(* IEC 61131-3 sources: SortJet_MasterSPS_Aufbau.fbsproj/Device.device.xml.v3^/Plc Logic.plclogic.xml.v3^/Application.application.xml.v3^/00_Basis/StationBasisZuweisungen.prg.st^, 20 files *)

(* ---- M_AufrufeZuweisungen.meth.st ---- *)
(* METADATA
{
	"v3Meta": {
		"objectGuid": "6343c508-4884-483e-a331-d4339a485652"
	}
}
*)
METHOD M_AufrufeZuweisungen
VAR_INPUT
END_VAR
VAR
  wlIndex : WORD;
END_VAR

//-------------------------------------------------------------------------------------------------
// PARAMETER ZUWEISEN
//-------------------------------------------------------------------------------------------------

// Aufrufe der Zuweisungen
Zuweisung_101();
Zuweisung_102();
Zuweisung_151();
Zuweisung_152();
Zuweisung_201();
Zuweisung_202();
Zuweisung_203();
Zuweisung_204();
Zuweisung_205();
Zuweisung_206();
Zuweisung_207();
Zuweisung_208();

Zuweisung_301();
Zuweisung_302();
Zuweisung_303();
Zuweisung_304();
Zuweisung_305();

Zuweisung_401();

Zuweisung_501();
END_METHOD

(* ---- Zuweisung_101.act.st ---- *)
(* METADATA
{
	"v3Meta": {
		"objectGuid": "51c9bc00-b1a7-48c3-ab96-ac2ea4b83acf"
	}
}
*)
ACTION Zuweisung_101
// Zuweisung der MK's
starrShuttleBasisParameter[cSHUTTLE_101].stMKs REF= apgMKShuttle101;

// Antriebsparameter zuweisen
starrShuttleBasisParameter[cSHUTTLE_101].stAntriebsparameter.stGlastransport                   REF= apgInfoShuttle101Glastransport;
starrShuttleBasisParameter[cSHUTTLE_101].stAntriebsparameter.stGlastransportSlave              REF= apgInfoShuttle101GlastransportSlave;
starrShuttleBasisParameter[cSHUTTLE_101].stAntriebsparameter.stWandverstellung                 REF= apgInfoShuttle101Dickenverstellung;
starrShuttleBasisParameter[cSHUTTLE_101].stParameterStationskomponenten.stGlastransportShuttle REF= apgMKShuttle101Glastransport;
starrShuttleBasisParameter[cSHUTTLE_101].stParameterStationskomponenten.stKippen               REF= apgMKShuttle101Kippen;
starrShuttleBasisParameter[cSHUTTLE_101].stParameterStationskomponenten.stWandverstellung      REF= apgMKShutte101Scheibenfuehrung;

starrShuttleBasisParameter[cSHUTTLE_101].stAntriebsparameter.stQuerfahrt REF= apgInfoShuttle101Querfahrt;
starrShuttleBasisParameter[cSHUTTLE_101].stAntriebsparameter.stKippen    REF= apgInfoShuttle101Kippen;

// Greifer [Ausbaustufe stStationsAufbau.bGreifer]
starrShuttleBasisParameter[cSHUTTLE_101].stParameterStationskomponenten.stGreifer REF= apgMKShuttle101Greifer;
starrShuttleBasisParameter[cSHUTTLE_101].stAntriebsparameter.stGreifer            REF= apgInfoShuttle101Greifer;

starrShuttleBasisParameter[cSHUTTLE_101].stParameterStationskomponenten.stZentralSchmierung REF= apgMKShuttleZentralschmierung[cSHUTTLE_101];

(* Hinweis:
   - Zuweisung der Transportrichtungen im Automatik-Betrieb für die Glastransporte
   - Zuweisungen der Kipp-Stati für die Übernahme/Übergabe an/von der jeweiligen Station
*)

// Transfershuttle des dynamischen Speichers  zuweisen
FOR wlIndex := cERSTES_TRANSFERSHUTTLE TO cLETZTES_TRANSFERSHUTTLE DO
  starrShuttleBasisParameter[cSHUTTLE_101].stMKs.stSchnittstellendaten.aEintransporte.Station[wlIndex]                  := Rueckwaertig;
  starrShuttleBasisParameter[cSHUTTLE_101].stMKs.stSchnittstellendaten.aEintransporte.Glastransport[wlIndex]            := eGlastransport_Default;
  starrShuttleBasisParameter[cSHUTTLE_101].stMKs.stSchnittstellendaten.aEintransporte.Kippen[wlIndex]                   := eKippen_Position_90Grad;
  starrShuttleBasisParameter[cSHUTTLE_101].stMKs.stSchnittstellendaten.aEintransporte.KippenNachEintransport[wlIndex]   := eKippen_Position_90Grad;
  starrShuttleBasisParameter[cSHUTTLE_101].stMKs.stSchnittstellendaten.aEintransporte.bStationQuittiertScheibe[wlIndex] := TRUE;

  starrShuttleBasisParameter[cSHUTTLE_101].stMKs.stSchnittstellendaten.aAustransporte.Station[wlIndex]                  := Vorwaertig;
  starrShuttleBasisParameter[cSHUTTLE_101].stMKs.stSchnittstellendaten.aAustransporte.Glastransport[wlIndex]            := eGlastransport_AufAuslauf;
  starrShuttleBasisParameter[cSHUTTLE_101].stMKs.stSchnittstellendaten.aAustransporte.Kippen[wlIndex]                   := eKippen_Position_90Grad;
  starrShuttleBasisParameter[cSHUTTLE_101].stMKs.stSchnittstellendaten.aAustransporte.KippenNachAustransport[wlIndex]   := eKippen_Position_84Grad;
  starrShuttleBasisParameter[cSHUTTLE_101].stMKs.stSchnittstellendaten.aAustransporte.bStationQuittiertScheibe[wlIndex] := TRUE;
END_FOR

// Station 207
starrShuttleBasisParameter[cSHUTTLE_101].stMKs.stSchnittstellendaten.aEintransporte.Station[cSTATION_207]                  := Rueckwaertig;
starrShuttleBasisParameter[cSHUTTLE_101].stMKs.stSchnittstellendaten.aEintransporte.Glastransport[cSTATION_207]            := eGlastransport_AufAuslaufVorab;
starrShuttleBasisParameter[cSHUTTLE_101].stMKs.stSchnittstellendaten.aEintransporte.Kippen[cSTATION_207]                   := eKippen_Position_90Grad;
starrShuttleBasisParameter[cSHUTTLE_101].stMKs.stSchnittstellendaten.aEintransporte.KippenNachEintransport[cSTATION_207]   := eKippen_Position_90Grad;
starrShuttleBasisParameter[cSHUTTLE_101].stMKs.stSchnittstellendaten.aEintransporte.bStationQuittiertScheibe[cSTATION_207] := TRUE;
END_ACTION

(* ---- Zuweisung_102.act.st ---- *)
(* METADATA
{
	"v3Meta": {
		"objectGuid": "58331703-c161-4204-81e2-c1518bdd5c02"
	}
}
*)
ACTION Zuweisung_102
// Zuweisung der MK's
starrShuttleBasisParameter[cSHUTTLE_102].stMKs REF= apgMKShuttle102;

// Antriebsparameter zuweisen
starrShuttleBasisParameter[cSHUTTLE_102].stAntriebsparameter.stGlastransport                   REF= apgInfoShuttle102Glastransport;
starrShuttleBasisParameter[cSHUTTLE_102].stAntriebsparameter.stGlastransportSlave              REF= apgInfoShuttle102GlastransportSlave;
starrShuttleBasisParameter[cSHUTTLE_102].stAntriebsparameter.stWandverstellung                 REF= apgInfoShuttle102Dickenverstellung;
starrShuttleBasisParameter[cSHUTTLE_102].stParameterStationskomponenten.stGlastransportShuttle REF= apgMKShuttle102Glastransport;
starrShuttleBasisParameter[cSHUTTLE_102].stParameterStationskomponenten.stKippen               REF= apgMKShuttle102Kippen;
starrShuttleBasisParameter[cSHUTTLE_102].stParameterStationskomponenten.stWandverstellung      REF= apgMKShutte102Scheibenfuehrung;

starrShuttleBasisParameter[cSHUTTLE_102].stAntriebsparameter.stQuerfahrt REF= apgInfoShuttle102Querfahrt;
starrShuttleBasisParameter[cSHUTTLE_102].stAntriebsparameter.stKippen    REF= apgInfoShuttle102Kippen;

// Greifer [Ausbaustufe stStationsAufbau.bGreifer]
starrShuttleBasisParameter[cSHUTTLE_102].stParameterStationskomponenten.stGreifer REF= apgMKShuttle102Greifer;
starrShuttleBasisParameter[cSHUTTLE_102].stAntriebsparameter.stGreifer            REF= apgInfoShuttle102Greifer;

starrShuttleBasisParameter[cSHUTTLE_102].stParameterStationskomponenten.stZentralSchmierung REF= apgMKShuttleZentralschmierung[cSHUTTLE_102];

(* Hinweis:
   - Zuweisung der Transportrichtungen im Automatik-Betrieb für die Glastransporte
   - Zuweisungen der Kipp-Stati für die Übernahme/Übergabe an/von der jeweiligen Station
*)

// Transfershuttle des dynamischen Speichers  zuweisen
FOR wlIndex := cERSTES_TRANSFERSHUTTLE TO cLETZTES_TRANSFERSHUTTLE DO
  starrShuttleBasisParameter[cSHUTTLE_102].stMKs.stSchnittstellendaten.aEintransporte.Station[wlIndex]                  := Vorwaertig;
  starrShuttleBasisParameter[cSHUTTLE_102].stMKs.stSchnittstellendaten.aEintransporte.Glastransport[wlIndex]            := eGlastransport_AufAuslauf;
  starrShuttleBasisParameter[cSHUTTLE_102].stMKs.stSchnittstellendaten.aEintransporte.Kippen[wlIndex]                   := eKippen_Position_90Grad;
  starrShuttleBasisParameter[cSHUTTLE_102].stMKs.stSchnittstellendaten.aEintransporte.KippenNachEintransport[wlIndex]   := eKippen_Position_90Grad;
  starrShuttleBasisParameter[cSHUTTLE_102].stMKs.stSchnittstellendaten.aEintransporte.bStationQuittiertScheibe[wlIndex] := TRUE;

  starrShuttleBasisParameter[cSHUTTLE_102].stMKs.stSchnittstellendaten.aAustransporte.Station[wlIndex]                  := Rueckwaertig;
  starrShuttleBasisParameter[cSHUTTLE_102].stMKs.stSchnittstellendaten.aAustransporte.Glastransport[wlIndex]            := eGlastransport_AufEinlaufVorab;
  starrShuttleBasisParameter[cSHUTTLE_102].stMKs.stSchnittstellendaten.aAustransporte.Kippen[wlIndex]                   := eKippen_Position_90Grad;
  starrShuttleBasisParameter[cSHUTTLE_102].stMKs.stSchnittstellendaten.aAustransporte.KippenNachAustransport[wlIndex]   := eKippen_Position_84Grad;
  starrShuttleBasisParameter[cSHUTTLE_102].stMKs.stSchnittstellendaten.aAustransporte.bStationQuittiertScheibe[wlIndex] := TRUE;
END_FOR

// Faecherwagenstationen: Austransport mit dem Greifer auf der Auslaufseite
FOR wlIndex := cERSTE_FAECHERWAGENSTATIONS_NR TO cLETZTE_FAECHERWAGENSTATIONS_NR DO
  starrShuttleBasisParameter[cSHUTTLE_102].stMKs.stSchnittstellendaten.aAustransporte.Station[wlIndex]                  := Vorwaertig;
  starrShuttleBasisParameter[cSHUTTLE_102].stMKs.stSchnittstellendaten.aAustransporte.Glastransport[wlIndex]            := eGlastransport_AufAuslauf;
  starrShuttleBasisParameter[cSHUTTLE_102].stMKs.stSchnittstellendaten.aAustransporte.Greifer[wlIndex]                  := eGreiferAuslaufseite;
  starrShuttleBasisParameter[cSHUTTLE_102].stMKs.stSchnittstellendaten.aAustransporte.bStationQuittiertScheibe[wlIndex] := TRUE;
END_FOR
END_ACTION

(* ---- Zuweisung_151.act.st ---- *)
(* METADATA
{
	"v3Meta": {
		"objectGuid": "626f2663-471d-49fb-b0f4-9d1f3bb0bf7f"
	}
}
*)
ACTION Zuweisung_151
// Zuweisung der MK's
starrTransfershuttleBasisParameter[cSHUTTLE_151].stMKs REF= apgMKTransfershuttle151;

// Antriebsparameter zuweisen
starrTransfershuttleBasisParameter[cSHUTTLE_151].stAntriebsparameter.stQuerfahrt             REF= apgInfoTransfershuttle151Querfahrt;
starrTransfershuttleBasisParameter[cSHUTTLE_151].stAntriebsparameter.stGlastransport         REF= apgInfoTransfer151Glastransport;

// Parameter der Stationskomponenten zuweisen
starrTransfershuttleBasisParameter[cSHUTTLE_151].stParameterStationskomponenten.stGlastransportTransferShuttle    REF= apgTransfer151Glastransport;
starrTransfershuttleBasisParameter[cSHUTTLE_151].stParameterStationskomponenten.stZentralSchmierung               REF= apgMKTransfershuttleZentralschmierung[cSHUTTLE_151];

(* Hinweis:
   - Zuweisung der Transportrichtungen im Automatik-Betrieb für die Glastransporte
   - Zuweisungen der Kipp-Stati für die Übernahme/Übergabe an/von der jeweiligen Station
*)
// Shuttle 101
starrTransfershuttleBasisParameter[cSHUTTLE_151].stMKs.stSchnittstellendaten.aEintransporte.Station[cSHUTTLE_101] := Vorwaertig;
starrTransfershuttleBasisParameter[cSHUTTLE_151].stMKs.stSchnittstellendaten.aAustransporte.Station[cSHUTTLE_101] := Rueckwaertig;

// Shuttle 102
starrTransfershuttleBasisParameter[cSHUTTLE_151].stMKs.stSchnittstellendaten.aEintransporte.Station[cSHUTTLE_102] := Rueckwaertig;
starrTransfershuttleBasisParameter[cSHUTTLE_151].stMKs.stSchnittstellendaten.aAustransporte.Station[cSHUTTLE_102] := Vorwaertig;
END_ACTION

(* ---- Zuweisung_152.act.st ---- *)
(* METADATA
{
	"v3Meta": {
		"objectGuid": "41f5393d-bf68-4ef4-aca8-1dae62f52119"
	}
}
*)
ACTION Zuweisung_152
// Zuweisung der MK's
starrTransfershuttleBasisParameter[cSHUTTLE_152].stMKs REF= apgMKTransfershuttle152;

// Antriebsparameter zuweisen
starrTransfershuttleBasisParameter[cSHUTTLE_152].stAntriebsparameter.stQuerfahrt             REF= apgInfoTransfershuttle152Querfahrt;
starrTransfershuttleBasisParameter[cSHUTTLE_152].stAntriebsparameter.stGlastransport         REF= apgInfoTransfer152Glastransport;

// Parameter der Stationskomponenten zuweisen
starrTransfershuttleBasisParameter[cSHUTTLE_152].stParameterStationskomponenten.stGlastransportTransferShuttle    REF= apgTransfer152Glastransport;
starrTransfershuttleBasisParameter[cSHUTTLE_152].stParameterStationskomponenten.stZentralSchmierung               REF= apgMKTransfershuttleZentralschmierung[cSHUTTLE_152];

(* Hinweis:
   - Zuweisung der Transportrichtungen im Automatik-Betrieb für die Glastransporte
   - Zuweisungen der Kipp-Stati für die Übernahme/Übergabe an/von der jeweiligen Station
*)
// Shuttle 101
starrTransfershuttleBasisParameter[cSHUTTLE_152].stMKs.stSchnittstellendaten.aEintransporte.Station[cSHUTTLE_101] := Vorwaertig;
starrTransfershuttleBasisParameter[cSHUTTLE_152].stMKs.stSchnittstellendaten.aAustransporte.Station[cSHUTTLE_101] := Rueckwaertig;

// Shuttle 102
starrTransfershuttleBasisParameter[cSHUTTLE_152].stMKs.stSchnittstellendaten.aEintransporte.Station[cSHUTTLE_102] := Rueckwaertig;
starrTransfershuttleBasisParameter[cSHUTTLE_152].stMKs.stSchnittstellendaten.aAustransporte.Station[cSHUTTLE_102] := Vorwaertig;
END_ACTION

(* ---- Zuweisung_201.act.st ---- *)
(* METADATA
{
	"v3Meta": {
		"objectGuid": "0d6757e1-53e1-48aa-88ce-f4bfba7d69cc"
	}
}
*)
ACTION Zuweisung_201
// Zuweisung der MK's
starrStationBasisParameter[cSTATION_201].stMKs REF= apgMKStation201;

// Antriebsparameter zuweisen
starrStationBasisParameter[cSTATION_201].stAntriebsparameter.stGlastransport         REF= apgInfoStation201Glastransport;
starrStationBasisParameter[cSTATION_201].stAntriebsparameter.stGlastransportSlave    REF= apgInfoStation201Glastransport_Slave;
starrStationBasisParameter[cSTATION_201].stAntriebsparameter.stMessachse             REF= apgInfoStation201Messachse;

// Parameter der Stationskomponenten zuweisen
starrStationBasisParameter[cSTATION_201].stParameterStationskomponenten.stGlastransport    REF= apgMKStation201Glastransport;
starrStationBasisParameter[cSTATION_201].stParameterStationskomponenten.stMessachse        REF= apgMKStation201Messachse;

(* Hinweis:
   - Zuweisung der Transportrichtungen im Automatik-Betrieb für die Glastransporte
   - Zuweisungen der Kipp-Stati für die Übernahme/Übergabe an/von der jeweiligen Station
*)

// Austransport
starrStationBasisParameter[cSTATION_201].stMKs.stSchnittstellendaten.aAustransporte.Station[cSTATION_202]                  := Vorwaertig;
starrStationBasisParameter[cSTATION_201].stMKs.stSchnittstellendaten.aAustransporte.bStationQuittiertScheibe[cSTATION_202] := FALSE;
END_ACTION

(* ---- Zuweisung_202.act.st ---- *)
(* METADATA
{
	"v3Meta": {
		"objectGuid": "e5688ce9-ab5a-4deb-8339-ae5087cb81c6"
	}
}
*)
ACTION Zuweisung_202
// Zuweisung der MK's
starrStationBasisParameter[cSTATION_202].stMKs REF= apgMKStation202;

// Antriebsparameter zuweisen
starrStationBasisParameter[cSTATION_202].stAntriebsparameter.stGlastransport               REF= apgInfoStation202Glastransport;
starrStationBasisParameter[cSTATION_202].stAntriebsparameter.stGlastransportSlave          REF= apgInfoStation202Glastransport_Slave;
starrStationBasisParameter[cSTATION_202].stAntriebsparameter.stKippen                      REF= apgInfoStation202Kippen;
starrStationBasisParameter[cSTATION_202].stAntriebsparameter.stQuerfahrt                   REF= apgInfoStation202Querfahrt;

// Parameter der Stationskomponenten zuweisen
starrStationBasisParameter[cSTATION_202].stParameterStationskomponenten.stGlastransport    REF= apgMKStation202Glastransport;
starrStationBasisParameter[cSTATION_202].stParameterStationskomponenten.stKippen           REF= apgMKStation202Kippen;
starrStationBasisParameter[cSTATION_202].stParameterStationskomponenten.stQuerfahrt        REF= apgMKStation202Querfahrt;

(* Hinweis:
   - Zuweisung der Transportrichtungen im Automatik-Betrieb für die Glastransporte
   - Zuweisungen der Kipp-Stati für die Übernahme/Übergabe an/von der jeweiligen Station
*)

// Eintransport
starrStationBasisParameter[cSTATION_202].stMKs.stSchnittstellendaten.aEintransporte.Station[cSTATION_201]                  := Vorwaertig;
starrStationBasisParameter[cSTATION_202].stMKs.stSchnittstellendaten.aEintransporte.Glastransport[cSTATION_201]            := eGlastransport_AufAuslaufVorab;
starrStationBasisParameter[cSTATION_202].stMKs.stSchnittstellendaten.aEintransporte.bStationQuittiertScheibe[cSTATION_201] := TRUE;

// Austransport
starrStationBasisParameter[cSTATION_202].stMKs.stSchnittstellendaten.aAustransporte.Station[cSTATION_203]                  := Vorwaertig;
starrStationBasisParameter[cSTATION_202].stMKs.stSchnittstellendaten.aAustransporte.bStationQuittiertScheibe[cSTATION_203] := FALSE;
END_ACTION

(* ---- Zuweisung_203.act.st ---- *)
(* METADATA
{
	"v3Meta": {
		"objectGuid": "120a0490-dc9c-46f0-83eb-c4f1579e8cf5"
	}
}
*)
ACTION Zuweisung_203
// Zuweisung der MK's
starrStationBasisParameter[cSTATION_203].stMKs REF= apgMKStation203;

// Antriebsparameter zuweisen
starrStationBasisParameter[cSTATION_203].stAntriebsparameter.stGlastransport               REF= apgInfoStation203Glastransport;
starrStationBasisParameter[cSTATION_203].stAntriebsparameter.stGlastransportSlave          REF= apgInfoStation203Glastransport_Slave;
starrStationBasisParameter[cSTATION_203].stAntriebsparameter.stKippen                      REF= apgInfoStation203Kippen;
starrStationBasisParameter[cSTATION_203].stAntriebsparameter.stQuerfahrt                   REF= apgInfoStation203Querfahrt;

// Parameter der Stationskomponenten zuweisen
starrStationBasisParameter[cSTATION_203].stParameterStationskomponenten.stGlastransport    REF= apgMKStation203Glastransport;
starrStationBasisParameter[cSTATION_203].stParameterStationskomponenten.stKippen           REF= apgMKStation203Kippen;
starrStationBasisParameter[cSTATION_203].stParameterStationskomponenten.stQuerfahrt        REF= apgMKStation203Querfahrt;

(* Hinweis:
   - Zuweisung der Transportrichtungen im Automatik-Betrieb für die Glastransporte
   - Zuweisungen der Kipp-Stati für die Übernahme/Übergabe an/von der jeweiligen Station
*)
// Eintransport
starrStationBasisParameter[cSTATION_203].stMKs.stSchnittstellendaten.aEintransporte.Station[cSTATION_202]                  := Vorwaertig;
starrStationBasisParameter[cSTATION_203].stMKs.stSchnittstellendaten.aEintransporte.Glastransport[cSTATION_202]            := eGlastransport_AufAuslaufVorab;
starrStationBasisParameter[cSTATION_203].stMKs.stSchnittstellendaten.aEintransporte.bStationQuittiertScheibe[cSTATION_202] := TRUE;

// Austransport
starrStationBasisParameter[cSTATION_203].stMKs.stSchnittstellendaten.aAustransporte.Station[cSTATION_204]                  := Vorwaertig;
starrStationBasisParameter[cSTATION_203].stMKs.stSchnittstellendaten.aAustransporte.bStationQuittiertScheibe[cSTATION_204] := FALSE;
END_ACTION

(* ---- Zuweisung_204.act.st ---- *)
(* METADATA
{
	"v3Meta": {
		"objectGuid": "508223db-73a6-4fc3-902d-ab2988c6447f"
	}
}
*)
ACTION Zuweisung_204
// Zuweisung der MK's
starrStationBasisParameter[cSTATION_204].stMKs REF= apgMKStation204;

// Antriebsparameter zuweisen
starrStationBasisParameter[cSTATION_204].stAntriebsparameter.stGlastransport             REF= apgInfoStation204Glastransport;
starrStationBasisParameter[cSTATION_204].stAntriebsparameter.stGlastransportSlave        REF= apgInfoStation204Glastransport_Slave;
starrStationBasisParameter[cSTATION_204].stAntriebsparameter.stGlastransportY            REF= apgInfoStation204GlastransportY;
starrStationBasisParameter[cSTATION_204].stAntriebsparameter.stGlastransportYSlave       REF= apgInfoStation204GlastransportY_Slave;

// Parameter der Stationskomponenten zuweisen
starrStationBasisParameter[cSTATION_204].stParameterStationskomponenten.stGlastransport  REF= apgMKStation204Glastransport;
starrStationBasisParameter[cSTATION_204].stParameterStationskomponenten.stGlastransportY REF= apgMKStation204GlastransportY;

// Hinweis:
// - Zuweisung der Transportrichtungen im Automatik-Betrieb fuer die Glastransporte
// - Achsrichtung: ueber welche Achse der Eckuebergabe mit der Nachbarstation transportiert wird

// Eintransport
starrStationBasisParameter[cSTATION_204].stMKs.stSchnittstellendaten.aEintransporte.Station[cSTATION_203]                  := Vorwaertig;
starrStationBasisParameter[cSTATION_204].stMKs.stSchnittstellendaten.aEintransporte.Glastransport[cSTATION_203]            := eGlastransport_AufAuslaufVorab;
starrStationBasisParameter[cSTATION_204].stMKs.stSchnittstellendaten.aEintransporte.Achsrichtung[cSTATION_203]             := eAchsrichtung_X;
starrStationBasisParameter[cSTATION_204].stMKs.stSchnittstellendaten.aEintransporte.bStationQuittiertScheibe[cSTATION_203] := TRUE;

starrStationBasisParameter[cSTATION_204].stMKs.stSchnittstellendaten.aEintransporte.Station[cSTATION_205]                  := Vorwaertig;
starrStationBasisParameter[cSTATION_204].stMKs.stSchnittstellendaten.aEintransporte.Glastransport[cSTATION_205]            := eGlastransport_AufAuslaufVorab;
starrStationBasisParameter[cSTATION_204].stMKs.stSchnittstellendaten.aEintransporte.Achsrichtung[cSTATION_205]             := eAchsrichtung_Y;
starrStationBasisParameter[cSTATION_204].stMKs.stSchnittstellendaten.aEintransporte.bStationQuittiertScheibe[cSTATION_205] := TRUE;

// Austransport
starrStationBasisParameter[cSTATION_204].stMKs.stSchnittstellendaten.aAustransporte.Station[cSTATION_206]                  := Vorwaertig;
starrStationBasisParameter[cSTATION_204].stMKs.stSchnittstellendaten.aAustransporte.Achsrichtung[cSTATION_206]             := eAchsrichtung_X;
starrStationBasisParameter[cSTATION_204].stMKs.stSchnittstellendaten.aAustransporte.bStationQuittiertScheibe[cSTATION_206] := FALSE;
END_ACTION

(* ---- Zuweisung_205.act.st ---- *)
(* METADATA
{
	"v3Meta": {
		"objectGuid": "e2d26e6b-cff2-4031-affb-248ab2534f79"
	}
}
*)
ACTION Zuweisung_205
// Zuweisung der MK's
starrStationBasisParameter[cSTATION_205].stMKs REF= apgMKStation205;

// Antriebsparameter zuweisen
starrStationBasisParameter[cSTATION_205].stAntriebsparameter.stGlastransport         REF= apgInfoStation205Glastransport;
starrStationBasisParameter[cSTATION_205].stAntriebsparameter.stGlastransportSlave    REF= apgInfoStation205Glastransport_Slave;
starrStationBasisParameter[cSTATION_205].stAntriebsparameter.stMessachse             REF= apgInfoStation205Messachse;

// Parameter der Stationskomponenten zuweisen
starrStationBasisParameter[cSTATION_205].stParameterStationskomponenten.stGlastransport    REF= apgMKStation205Glastransport;
starrStationBasisParameter[cSTATION_205].stParameterStationskomponenten.stMessachse        REF= apgMKStation205Messachse;

(* Hinweis:
   - Zuweisung der Transportrichtungen im Automatik-Betrieb für die Glastransporte
   - Zuweisungen der Kipp-Stati für die Übernahme/Übergabe an/von der jeweiligen Station
*)

// Eintransport
starrStationBasisParameter[cSTATION_205].stMKs.stSchnittstellendaten.aEintransporte.Station[cFREMDANLAGE_EINLAUF_1]                  := Vorwaertig;
starrStationBasisParameter[cSTATION_205].stMKs.stSchnittstellendaten.aEintransporte.Glastransport[cFREMDANLAGE_EINLAUF_1]            := eGlastransport_AufAuslaufVorab;
starrStationBasisParameter[cSTATION_205].stMKs.stSchnittstellendaten.aEintransporte.bStationQuittiertScheibe[cFREMDANLAGE_EINLAUF_1] := TRUE;

// Austransport
starrStationBasisParameter[cSTATION_205].stMKs.stSchnittstellendaten.aAustransporte.Station[cSTATION_204]                  := Vorwaertig;
starrStationBasisParameter[cSTATION_205].stMKs.stSchnittstellendaten.aAustransporte.bStationQuittiertScheibe[cSTATION_204] := FALSE;
END_ACTION

(* ---- Zuweisung_206.act.st ---- *)
(* METADATA
{
	"v3Meta": {
		"objectGuid": "ec549a81-8212-4c0f-885a-b7f66d397584"
	}
}
*)
ACTION Zuweisung_206
// Zuweisung der MK's
starrStationBasisParameter[cSTATION_206].stMKs REF= apgMKStation206;

// Antriebsparameter zuweisen
starrStationBasisParameter[cSTATION_206].stAntriebsparameter.stGlastransport               REF= apgInfoStation206Glastransport;
starrStationBasisParameter[cSTATION_206].stAntriebsparameter.stGlastransportSlave          REF= apgInfoStation206Glastransport_Slave;
starrStationBasisParameter[cSTATION_206].stAntriebsparameter.stQuerfahrt                   REF= apgInfoStation206Querfahrt;
starrStationBasisParameter[cSTATION_206].stAntriebsparameter.stKippen                      REF= apgInfoStation206Kippen;

// Parameter der Stationskomponenten zuweisen
starrStationBasisParameter[cSTATION_206].stParameterStationskomponenten.stGlastransport    REF= apgMKStation206Glastransport;
starrStationBasisParameter[cSTATION_206].stParameterStationskomponenten.stQuerfahrt        REF= apgMKStation206Querfahrt;
starrStationBasisParameter[cSTATION_206].stParameterStationskomponenten.stKippen           REF= apgMKStation206Kippen;

(* Hinweis:
   - Zuweisung der Transportrichtungen im Automatik-Betrieb für die Glastransporte
   - Zuweisungen der Kipp-Stati für die Übernahme/Übergabe an/von der jeweiligen Station
*)

// Eintransport von der Eckuebergabe 204
starrStationBasisParameter[cSTATION_206].stMKs.stSchnittstellendaten.aEintransporte.Station[cSTATION_204]                  := Vorwaertig;
starrStationBasisParameter[cSTATION_206].stMKs.stSchnittstellendaten.aEintransporte.Glastransport[cSTATION_204]            := eGlastransport_AufAuslaufVorab;
starrStationBasisParameter[cSTATION_206].stMKs.stSchnittstellendaten.aEintransporte.Kippen[cSTATION_204]                   := eKippen_Position_0Grad;
starrStationBasisParameter[cSTATION_206].stMKs.stSchnittstellendaten.aEintransporte.KippenNachEintransport[cSTATION_204]   := eKippen_Position_84Grad;
starrStationBasisParameter[cSTATION_206].stMKs.stSchnittstellendaten.aEintransporte.bStationQuittiertScheibe[cSTATION_204] := TRUE;

// Austransport an die Drehstation 207
starrStationBasisParameter[cSTATION_206].stMKs.stSchnittstellendaten.aAustransporte.Station[cSTATION_207]                  := Vorwaertig;
starrStationBasisParameter[cSTATION_206].stMKs.stSchnittstellendaten.aAustransporte.Kippen[cSTATION_207]                   := eKippen_Position_84Grad;
starrStationBasisParameter[cSTATION_206].stMKs.stSchnittstellendaten.aAustransporte.KippenNachAustransport[cSTATION_207]   := eKippen_Position_0Grad;
starrStationBasisParameter[cSTATION_206].stMKs.stSchnittstellendaten.aAustransporte.bStationQuittiertScheibe[cSTATION_207] := FALSE;
END_ACTION

(* ---- Zuweisung_207.act.st ---- *)
(* METADATA
{
	"v3Meta": {
		"objectGuid": "f55699bd-423e-450f-9568-477ca85fd454"
	}
}
*)
ACTION Zuweisung_207
// Zuweisung der MK's
starrStationBasisParameter[cSTATION_207].stMKs REF= apgMKStation207;

// Antriebsparameter zuweisen
starrStationBasisParameter[cSTATION_207].stAntriebsparameter.stGlastransport            REF= apgInfoStation207Glastransport;
starrStationBasisParameter[cSTATION_207].stAntriebsparameter.stGlastransportSlave       REF= apgInfoStation207GlastransportSlave;
starrStationBasisParameter[cSTATION_207].stAntriebsparameter.stDrehen                   REF= apgInfoStation207Drehen;
starrStationBasisParameter[cSTATION_207].stAntriebsparameter.stKippen                   REF= apgInfoStation207Kippen;
starrStationBasisParameter[cSTATION_207].stAntriebsparameter.stQuerfahrt                REF= apgInfoStation207Querfahrt;

// Parameter der Stationskomponenten zuweisen
starrStationBasisParameter[cSTATION_207].stParameterStationskomponenten.stGlastransport REF= apgMKStation207Glastransport;
starrStationBasisParameter[cSTATION_207].stParameterStationskomponenten.stDrehen        REF= apgMKStation207Drehen;
starrStationBasisParameter[cSTATION_207].stParameterStationskomponenten.stKippen        REF= apgMKStation207Kippen;
starrStationBasisParameter[cSTATION_207].stParameterStationskomponenten.stQuerfahrt     REF= apgMKStation207Querfahrt;

(* Hinweis:
   - Zuweisung der Transportrichtungen im Automatik-Betrieb für die Glastransporte
   - Drehpositionen der Drehstation:
       90 Grad      -> Anlegewand 208
       0 / 180 Grad -> Kipptisch 206 / Shuttle 101 (0 Grad = bisherige 90-Grad-Position, 180 Grad = um 180 Grad gedreht)
   - Drehpositionen kommen aktuell aus dieser Zuweisung (MK bDrehpositionenVomMMI = FALSE): Drehen / DrehenNachEintransport /
     DrehenNachAustransport unten gelten. Spaeter kommen sie vom MMI (bDrehpositionenVomMMI = TRUE), dann werden die
     Drehen-Eintraege hier nicht mehr ausgewertet.
   - Kippen der Drehstation VOR der Aktion kommt aus den Kippen-Eintraegen hier (Kippen),
     NACH dem Ein- und Austransport aus KippenNachEintransport / KippenNachAustransport.
     Nur der Systemcheck nimmt die Kippposition aus der Drehposition (MK: apgMKStation207Drehen.astKippenJeDrehposition).
*)

// Eintransport von der Anlegewand 208 (Drehposition 90 Grad, vom MMI)
starrStationBasisParameter[cSTATION_207].stMKs.stSchnittstellendaten.aEintransporte.Station[cSTATION_208]                  := Rueckwaertig;
starrStationBasisParameter[cSTATION_207].stMKs.stSchnittstellendaten.aEintransporte.Glastransport[cSTATION_208]            := eGlastransport_AufAuslaufVorab;
starrStationBasisParameter[cSTATION_207].stMKs.stSchnittstellendaten.aEintransporte.Kippen[cSTATION_208]                   := eKippen_Position_84Grad;
starrStationBasisParameter[cSTATION_207].stMKs.stSchnittstellendaten.aEintransporte.KippenNachEintransport[cSTATION_208]   := eKippen_Position_90Grad;
starrStationBasisParameter[cSTATION_207].stMKs.stSchnittstellendaten.aEintransporte.Drehen[cSTATION_208]                   := eDrehPosition90Grad;
starrStationBasisParameter[cSTATION_207].stMKs.stSchnittstellendaten.aEintransporte.DrehenNachEintransport[cSTATION_208]   := eDrehPosition0Grad;
starrStationBasisParameter[cSTATION_207].stMKs.stSchnittstellendaten.aEintransporte.bStationQuittiertScheibe[cSTATION_208] := TRUE;

// Eintransport vom Kipptisch 206 (Drehposition 0 / 180 Grad, vom MMI)
starrStationBasisParameter[cSTATION_207].stMKs.stSchnittstellendaten.aEintransporte.Station[cSTATION_206]                  := Vorwaertig;
starrStationBasisParameter[cSTATION_207].stMKs.stSchnittstellendaten.aEintransporte.Glastransport[cSTATION_206]            := eGlastransport_AufAuslaufVorab;
starrStationBasisParameter[cSTATION_207].stMKs.stSchnittstellendaten.aEintransporte.Kippen[cSTATION_206]                   := eKippen_Position_84Grad;
starrStationBasisParameter[cSTATION_207].stMKs.stSchnittstellendaten.aEintransporte.KippenNachEintransport[cSTATION_206]   := eKippen_Position_90Grad;
starrStationBasisParameter[cSTATION_207].stMKs.stSchnittstellendaten.aEintransporte.Drehen[cSTATION_206]                   := eDrehPosition0Grad;
starrStationBasisParameter[cSTATION_207].stMKs.stSchnittstellendaten.aEintransporte.DrehenNachEintransport[cSTATION_206]   := eDrehPosition0Grad;
starrStationBasisParameter[cSTATION_207].stMKs.stSchnittstellendaten.aEintransporte.bStationQuittiertScheibe[cSTATION_206] := TRUE;

// Austransport an das Shuttle 101 (Drehposition 0 / 180 Grad, vom MMI)
starrStationBasisParameter[cSTATION_207].stMKs.stSchnittstellendaten.aAustransporte.Station[cSHUTTLE_101]                  := Vorwaertig;
starrStationBasisParameter[cSTATION_207].stMKs.stSchnittstellendaten.aAustransporte.Kippen[cSHUTTLE_101]                   := eKippen_Position_90Grad;
starrStationBasisParameter[cSTATION_207].stMKs.stSchnittstellendaten.aAustransporte.KippenNachAustransport[cSHUTTLE_101]   := eKippen_Position_84Grad;
starrStationBasisParameter[cSTATION_207].stMKs.stSchnittstellendaten.aAustransporte.Drehen[cSHUTTLE_101]                   := eDrehPosition0Grad;
starrStationBasisParameter[cSTATION_207].stMKs.stSchnittstellendaten.aAustransporte.DrehenNachAustransport[cSHUTTLE_101]   := eDrehPosition0Grad;
starrStationBasisParameter[cSTATION_207].stMKs.stSchnittstellendaten.aAustransporte.bStationQuittiertScheibe[cSHUTTLE_101] := FALSE;
END_ACTION

(* ---- Zuweisung_208.act.st ---- *)
(* METADATA
{
	"v3Meta": {
		"objectGuid": "c063edf5-417b-4a06-b1eb-b2a6b64450cf"
	}
}
*)
ACTION Zuweisung_208
// Zuweisung der MK's
starrStationBasisParameter[cSTATION_208].stMKs REF= apgMKStation208;

// Antriebsparameter zuweisen
starrStationBasisParameter[cSTATION_208].stAntriebsparameter.stGlastransport               REF= apgInfoStation208Glastransport;
starrStationBasisParameter[cSTATION_208].stAntriebsparameter.stGlastransportSlave          REF= apgInfoStation208GlastransportSlave;
starrStationBasisParameter[cSTATION_208].stAntriebsparameter.stMessachse                   REF= apgInfoStation208Messachse;
starrStationBasisParameter[cSTATION_208].stAntriebsparameter.stKippen                      REF= apgInfoStation208Kippen;

// Parameter der Stationskomponenten zuweisen
starrStationBasisParameter[cSTATION_208].stParameterStationskomponenten.stGlastransport    REF= apgMKStation208Glastransport;
starrStationBasisParameter[cSTATION_208].stParameterStationskomponenten.stMessachse        REF= apgMKStation208Messachse;
starrStationBasisParameter[cSTATION_208].stParameterStationskomponenten.stKippen           REF= apgMKStation208Kippen;

(* Hinweis:
   - Zuweisung der Transportrichtungen im Automatik-Betrieb für die Glastransporte
   - Zuweisungen der Kipp-Stati für die Übernahme/Übergabe an/von der jeweiligen Station
*)

// Eintransport
// Nicht vorhanden

// Austransport
starrStationBasisParameter[cSTATION_208].stMKs.stSchnittstellendaten.aAustransporte.Station[cSTATION_207]                  := Vorwaertig;
starrStationBasisParameter[cSTATION_208].stMKs.stSchnittstellendaten.aAustransporte.bStationQuittiertScheibe[cSTATION_207] := FALSE;
END_ACTION

(* ---- Zuweisung_301.act.st ---- *)
(* METADATA
{
	"v3Meta": {
		"objectGuid": "f22c61c3-e14c-4dd4-a956-6cafd549323c"
	}
}
*)
ACTION Zuweisung_301
// Zuweisung der MK's
starrFaecherwagenBasisParameter[cSTATION_301].stMKs REF= apgMKFaecherwagenstation[cSTATION_301];

// Zuweisung Sammel-IOs
// in_bDruckluftOK: wird zyklisch beim Aufruf in StationsAufrufe (MainTask) uebergeben - nicht hier (SlowTask, Mehrfach-Task-Zugriff auf E/As)
END_ACTION

(* ---- Zuweisung_302.act.st ---- *)
(* METADATA
{
	"v3Meta": {
		"objectGuid": "bc82e65a-c6a0-47b9-a190-18e8260f866e"
	}
}
*)
ACTION Zuweisung_302
// Zuweisung der MK's
starrFaecherwagenBasisParameter[cSTATION_302].stMKs REF= apgMKFaecherwagenstation[cSTATION_302];

// Zuweisung Sammel-IOs
// in_bDruckluftOK: wird zyklisch beim Aufruf in StationsAufrufe (MainTask) uebergeben - nicht hier (SlowTask, Mehrfach-Task-Zugriff auf E/As)
END_ACTION

(* ---- Zuweisung_303.act.st ---- *)
(* METADATA
{
	"v3Meta": {
		"objectGuid": "150cb19f-2e3d-4826-8e12-7d1c3a1232ee"
	}
}
*)
ACTION Zuweisung_303
// Zuweisung der MK's
starrFaecherwagenBasisParameter[cSTATION_303].stMKs REF= apgMKFaecherwagenstation[cSTATION_303];

// Zuweisung Sammel-IOs
// in_bDruckluftOK: wird zyklisch beim Aufruf in StationsAufrufe (MainTask) uebergeben - nicht hier (SlowTask, Mehrfach-Task-Zugriff auf E/As)
END_ACTION

(* ---- Zuweisung_304.act.st ---- *)
(* METADATA
{
	"v3Meta": {
		"objectGuid": "50ec10ce-5886-414e-95bc-f0e33c3a8c61"
	}
}
*)
ACTION Zuweisung_304
// Zuweisung der MK's
starrFaecherwagenBasisParameter[cSTATION_304].stMKs REF= apgMKFaecherwagenstation[cSTATION_304];

// Zuweisung Sammel-IOs
// in_bDruckluftOK: wird zyklisch beim Aufruf in StationsAufrufe (MainTask) uebergeben - nicht hier (SlowTask, Mehrfach-Task-Zugriff auf E/As)
END_ACTION

(* ---- Zuweisung_305.act.st ---- *)
(* METADATA
{
	"v3Meta": {
		"objectGuid": "1eb663c8-b9f8-4b76-a432-de5bea4a687b"
	}
}
*)
ACTION Zuweisung_305
// Zuweisung der MK's
starrFaecherwagenBasisParameter[cSTATION_305].stMKs REF= apgMKFaecherwagenstation[cSTATION_305];

// Zuweisung Sammel-IOs
// in_bDruckluftOK: wird zyklisch beim Aufruf in StationsAufrufe (MainTask) uebergeben - nicht hier (SlowTask, Mehrfach-Task-Zugriff auf E/As)
END_ACTION

(* ---- Zuweisung_401.act.st ---- *)
(* METADATA
{
	"v3Meta": {
		"objectGuid": "4728ef0b-ed05-4ab8-920f-4f7ee6482110"
	}
}
*)
ACTION Zuweisung_401
// Zuweisung der MK's
starrFremdanlageAuslaufStationBasisParameter[cSTATION_401].stMKs REF= apgMKStation401;
END_ACTION

(* ---- Zuweisung_501.act.st ---- *)
(* METADATA
{
	"v3Meta": {
		"objectGuid": "ec9cfad2-6d06-4c52-981e-45ef0970cfa5"
	}
}
*)
ACTION Zuweisung_501
// Zuweisung der MK's
starrFremdanlageEinlaufStationBasisParameter[cFREMDANLAGE_EINLAUF_1].stMKs REF= apgMKStation501;
END_ACTION
